FUNCTION_BLOCK Draining
VAR_INPUT
	diEnabled : BOOL;
END_VAR
VAR_OUTPUT
	doEnabled : BOOL;
END_VAR
VAR_IN_OUT
	DrainingPhase : TPhaseDraining;
	DrainingValve : TValve;
END_VAR
VAR
END_VAR

{region "Aut/Man"}
    // switching state of engine - automatic or manual control (default state is manual)
    IF DrainingPhase.Cmd.AutCtrl AND NOT DrainingPhase.State.AutCtrl THEN
        DrainingPhase.State.AutCtrl := TRUE;
        DrainingPhase.State.ManCtrl := FALSE;
        DrainingPhase.State.Running := FALSE;
        DrainingPhase.State.Paused  := FALSE;
        DrainingPhase.State.Idle    := TRUE;
    ELSIF DrainingPhase.Cmd.ManCtrl AND NOT DrainingPhase.State.ManCtrl THEN
        DrainingPhase.State.ManCtrl := TRUE;
        DrainingPhase.State.AutCtrl := FALSE;
        DrainingPhase.State.Running := FALSE;
        DrainingPhase.State.Paused  := FALSE;
        DrainingPhase.State.Idle    := TRUE;
    END_IF;

    IF NOT DrainingPhase.State.AutCtrl AND NOT DrainingPhase.State.ManCtrl THEN
        DrainingPhase.State.ManCtrl := TRUE;
    END_IF;

    DrainingPhase.Cmd.AutCtrl := FALSE;
    DrainingPhase.Cmd.ManCtrl := FALSE;
{endregion}

{region "ManCtrl"}
    // processing manual actions - if command is processed, it is sets to FALSE even if can't be processed
    IF DrainingPhase.State.ManCtrl THEN

        // Start - open draining valve
        IF DrainingPhase.Cmd.StartMan AND DrainingPhase.State.Idle AND NOT DrainingValve.State.GenErr THEN
            DrainingPhase.State.Idle    := FALSE;
            DrainingPhase.State.Running := TRUE;
            DrainingPhase.State.Done    := FALSE;
            DrainingValve.Cmd.AutCtrl   := TRUE;   // valve must be in auto, the phase drives it by requests
        END_IF;
        // Stop - close draining valve
        IF DrainingPhase.Cmd.StopMan AND (DrainingPhase.State.Running OR DrainingPhase.State.Paused) THEN
            DrainingPhase.State.Running := FALSE;
            DrainingPhase.State.Paused  := FALSE;
            DrainingPhase.State.Idle    := TRUE;
        END_IF;
        // Pause - close draining valve
        IF DrainingPhase.Cmd.PauseMan AND DrainingPhase.State.Running THEN
            DrainingPhase.State.Running := FALSE;
            DrainingPhase.State.Paused  := TRUE;
        END_IF;
        // Resume - open draining valve
        IF DrainingPhase.Cmd.ResumeMan AND DrainingPhase.State.Paused AND NOT DrainingValve.State.GenErr THEN
            DrainingPhase.State.Paused  := FALSE;
            DrainingPhase.State.Running := TRUE;
        END_IF;
    // real states of phase are writed into states in phase structure
    END_IF;
    DrainingPhase.Cmd.StartMan  := FALSE;
    DrainingPhase.Cmd.StopMan   := FALSE;
    DrainingPhase.Cmd.PauseMan  := FALSE;
    DrainingPhase.Cmd.ResumeMan := FALSE;
{endregion}

{region "AutCtrl"}
    //if request to run in automatic mode -> set auto request to open of filling valve to 1 and close to 0, if not open 0 close 1
    IF DrainingPhase.State.AutCtrl THEN
        IF DrainingPhase.Cmd.StartAut AND DrainingPhase.State.Idle AND NOT DrainingValve.State.GenErr THEN
            DrainingPhase.State.Idle    := FALSE;
            DrainingPhase.State.Running := TRUE;
            DrainingPhase.State.Done    := FALSE;
            DrainingValve.Cmd.AutCtrl   := TRUE;
        END_IF;

        IF DrainingPhase.Cmd.StopAut AND (DrainingPhase.State.Running OR DrainingPhase.State.Paused) THEN
            DrainingPhase.State.Running := FALSE;
            DrainingPhase.State.Paused  := FALSE;
            DrainingPhase.State.Idle    := TRUE;
        END_IF;
    END_IF;
    // commands should be sets to false after their processing
    DrainingPhase.Cmd.StartAut := FALSE;
    DrainingPhase.Cmd.StopAut  := FALSE;
{endregion}
{region "Done"}
    //every phase should have finish condition - draining phase - if water level is below requested level
    //after that done state should be setted to 1
    IF DrainingPhase.State.Running AND (DrainingPhase.WaterLevel <= DrainingPhase.ParamDrainLevel) THEN
        DrainingPhase.State.Running := FALSE;
        DrainingPhase.State.Idle    := TRUE;
        DrainingPhase.State.Done    := TRUE;
    END_IF;
    IF DrainingPhase.Cmd.ResetDone THEN
        DrainingPhase.State.Done := FALSE;
        DrainingPhase.Cmd.ResetDone := FALSE;
    END_IF;
{endregion}

{region "States"} 
    //Command valve in cases of states
    IF DrainingPhase.State.Running AND DrainingValve.State.GenErr THEN
        DrainingPhase.State.Running := FALSE;
        DrainingPhase.State.Paused  := TRUE;
    END_IF;

    IF DrainingPhase.State.Running THEN
        DrainingValve.Cmd.Req2OpenAut  := TRUE;
        DrainingValve.Cmd.Req2CloseAut := FALSE;
    ELSE
        DrainingValve.Cmd.Req2OpenAut  := FALSE;
        DrainingValve.Cmd.Req2CloseAut := TRUE;
    END_IF;
{endregion}

// delault state of phase - if not any state sets state to idle
IF (NOT DrainingPhase.State.Idle) AND (NOT DrainingPhase.State.Paused) AND (NOT DrainingPhase.State.Running) THEN
    DrainingPhase.State.Idle := 1;
END_IF;

// write binary states into int value for visualization
IF DrainingPhase.State.Idle THEN
    DrainingPhase.State.StateInt := Global.PhIdle;
ELSIF DrainingPhase.State.Running THEN
    DrainingPhase.State.StateInt := Global.PhRunning;
ELSE
    DrainingPhase.State.StateInt := Global.PhPause;
END_IF;

//Ponechte pro moznost retezeni volani bloku v LAD
doEnabled := diEnabled;

END_FUNCTION_BLOCK

(* stored: Version 1.1.0.1, ProductVersion 3.1.4024.13
   POU Draining: Id {a501d01f-bc41-415b-8bb8-19a7a35d7bf8}, SpecialFunc None *)
